(* IEC 61131-3 sources: plc-st-coding-agent/progress/evidence/f14_v6_public_pilot_20261112/jobs/custom_minimax-m27, 44 files *)

(* ---- public-easy-01.candidate_01.st ---- *)
FUNCTION_BLOCK FillLineControl
VAR_INPUT
    bottleSensor           : BOOL;
    cleaningConfirmButton  : BOOL;
    fillingConfirmButton   : BOOL;
    cappingConfirmButton   : BOOL;
    packingConfirmButton   : BOOL;
    finishedButton         : BOOL;
END_VAR

VAR_OUTPUT
    Pump_Motor         : BOOL;
    Filling_Valve      : BOOL;
    Capping_Machine    : BOOL;
    Packing_Machine    : BOOL;
    Completion_Light   : BOOL;
END_VAR

VAR
    eState : INT;
    tmp_R_TRIG_cleaning : R_TRIG;
    tmp_R_TRIG_filling  : R_TRIG;
    tmp_R_TRIG_capping  : R_TRIG;
    tmp_R_TRIG_packing  : R_TRIG;
    tmp_R_TRIG_finished : R_TRIG;
END_VAR

VAR CONSTANT
    STATE_IDLE      : INT := 0;
    STATE_CLEANING  : INT := 1;
    STATE_FILLING   : INT := 2;
    STATE_CAPPING   : INT := 3;
    STATE_PACKING   : INT := 4;
    STATE_COMPLETED : INT := 5;
END_VAR

(* ENGINEERING_CONTRACT
  State machine for automated filling line (6 states, linear sequence):
  +------------------+-------------------------------+-------------------+-------------------+---------------------------+
  | State            | Active Outputs                | Retention         | Deactivation      | Trigger                   |
  +------------------+-------------------------------+-------------------+-------------------+---------------------------+
  | IDLE (0)         | none                          | N/A               | N/A               | bottleSensor=TRUE         |
  | CLEANING (1)     | Pump_Motor=TRUE               | Hold until next   | Next state enter  | cleaningConfirmButton edge|
  | FILLING (2)      | Filling_Valve=TRUE            | Hold until next   | Next state enter  | fillingConfirmButton edge |
  | CAPPING (3)      | Capping_Machine=TRUE          | Hold until next   | Next state enter  | cappingConfirmButton edge |
  | PACKING (4)      | Packing_Machine=TRUE          | Hold until next   | Next state enter  | packingConfirmButton edge |
  | COMPLETED (5)    | Completion_Light=TRUE         | Hold until reset  | finishedButton edge | packingConfirmButton edge|
  +------------------+-------------------------------+-------------------+-------------------+---------------------------+
  Priority: Same-scan parallel evaluation, outputs set per state at scan end.
  References: PUB003(cleaning pump start), PUB004(cleaningConfirmButton),
              PUB005(fillingConfirmButton), PUB006(cappingConfirmButton),
              PUB007(packingConfirmButton), PUB008(finishedButton reset).
*)
(* CONTRACT_RULES [{"kind":"hold_until_reset","output":"Completion_Light","set_input":"packingConfirmButton","reset_input":"finishedButton"}] *)

tmp_R_TRIG_cleaning(CLK := cleaningConfirmButton);
tmp_R_TRIG_filling(CLK  := fillingConfirmButton);
tmp_R_TRIG_capping(CLK  := cappingConfirmButton);
tmp_R_TRIG_packing(CLK  := packingConfirmButton);
tmp_R_TRIG_finished(CLK := finishedButton);

CASE eState OF
    STATE_IDLE:
        Pump_Motor       := FALSE;
        Filling_Valve    := FALSE;
        Capping_Machine  := FALSE;
        Packing_Machine  := FALSE;
        Completion_Light := FALSE;

        IF bottleSensor THEN
            eState := STATE_CLEANING;
        END_IF;

    STATE_CLEANING:
        Pump_Motor       := TRUE;
        Filling_Valve    := FALSE;
        Capping_Machine  := FALSE;
        Packing_Machine  := FALSE;
        Completion_Light := FALSE;

        IF tmp_R_TRIG_cleaning.Q THEN
            eState := STATE_FILLING;
        END_IF;

    STATE_FILLING:
        Pump_Motor       := FALSE;
        Filling_Valve    := TRUE;
        Capping_Machine  := FALSE;
        Packing_Machine  := FALSE;
        Completion_Light := FALSE;

        IF tmp_R_TRIG_filling.Q THEN
            eState := STATE_CAPPING;
        END_IF;

    STATE_CAPPING:
        Pump_Motor       := FALSE;
        Filling_Valve    := FALSE;
        Capping_Machine  := TRUE;
        Packing_Machine  := FALSE;
        Completion_Light := FALSE;

        IF tmp_R_TRIG_capping.Q THEN
            eState := STATE_PACKING;
        END_IF;

    STATE_PACKING:
        Pump_Motor       := FALSE;
        Filling_Valve    := FALSE;
        Capping_Machine  := FALSE;
        Packing_Machine  := TRUE;
        Completion_Light := FALSE;

        IF tmp_R_TRIG_packing.Q THEN
            eState := STATE_COMPLETED;
        END_IF;

    STATE_COMPLETED:
        Pump_Motor       := FALSE;
        Filling_Valve    := FALSE;
        Capping_Machine  := FALSE;
        Packing_Machine  := FALSE;
        Completion_Light := TRUE;

        IF tmp_R_TRIG_finished.Q THEN
            eState := STATE_IDLE;
        END_IF;
END_CASE;

END_FUNCTION_BLOCK

(* ---- public-easy-01.candidate_02.st ---- *)
FUNCTION_BLOCK FillLineControl
VAR_INPUT
    bottleSensor           : BOOL;
    cleaningConfirmButton  : BOOL;
    fillingConfirmButton   : BOOL;
    cappingConfirmButton   : BOOL;
    packingConfirmButton   : BOOL;
    finishedButton         : BOOL;
END_VAR

VAR_OUTPUT
    Pump_Motor         : BOOL;
    Filling_Valve      : BOOL;
    Capping_Machine    : BOOL;
    Packing_Machine    : BOOL;
    Completion_Light   : BOOL;
END_VAR

VAR
    eState : INT;
    tmp_R_TRIG_cleaning : R_TRIG;
    tmp_R_TRIG_filling  : R_TRIG;
    tmp_R_TRIG_capping  : R_TRIG;
    tmp_R_TRIG_packing  : R_TRIG;
    tmp_R_TRIG_finished : R_TRIG;
END_VAR

VAR CONSTANT
    STATE_IDLE      : INT := 0;
    STATE_CLEANING  : INT := 1;
    STATE_FILLING   : INT := 2;
    STATE_CAPPING   : INT := 3;
    STATE_PACKING   : INT := 4;
    STATE_COMPLETED : INT := 5;
END_VAR

(* ENGINEERING_CONTRACT
  State machine for automated filling line (6 states, linear sequence):
  +------------------+-------------------------------+-------------------+-------------------+---------------------------+
  | State            | Active Outputs                | Retention         | Deactivation      | Trigger                   |
  +------------------+-------------------------------+-------------------+-------------------+---------------------------+
  | IDLE (0)         | none                          | N/A               | N/A               | bottleSensor=TRUE         |
  | CLEANING (1)     | Pump_Motor=TRUE               | Hold until next   | Next state enter  | cleaningConfirmButton edge|
  | FILLING (2)      | Filling_Valve=TRUE            | Hold until next   | Next state enter  | fillingConfirmButton edge |
  | CAPPING (3)      | Capping_Machine=TRUE          | Hold until next   | Next state enter  | cappingConfirmButton edge |
  | PACKING (4)      | Packing_Machine=TRUE          | Hold until next   | Next state enter  | packingConfirmButton edge |
  | COMPLETED (5)    | Completion_Light=TRUE         | Hold until reset  | finishedButton edge | -                      |
  +------------------+-------------------------------+-------------------+-------------------+---------------------------+
  Priority: Same-scan parallel evaluation, outputs set per state at scan end.
  Completion_Light set_input (packingConfirmButton) requires reaching STATE_PACKING first;
  this prerequisite cannot be expressed in flat contract format and is handled by the
  state machine logic. PUB003-PUB008 define all transitions.
*)
(* CONTRACT_RULES [] *)

tmp_R_TRIG_cleaning(CLK := cleaningConfirmButton);
tmp_R_TRIG_filling(CLK  := fillingConfirmButton);
tmp_R_TRIG_capping(CLK  := cappingConfirmButton);
tmp_R_TRIG_packing(CLK  := packingConfirmButton);
tmp_R_TRIG_finished(CLK := finishedButton);

CASE eState OF
    STATE_IDLE:
        Pump_Motor       := FALSE;
        Filling_Valve    := FALSE;
        Capping_Machine  := FALSE;
        Packing_Machine  := FALSE;
        Completion_Light := FALSE;

        IF bottleSensor THEN
            eState := STATE_CLEANING;
        END_IF;

    STATE_CLEANING:
        Pump_Motor       := TRUE;
        Filling_Valve    := FALSE;
        Capping_Machine  := FALSE;
        Packing_Machine  := FALSE;
        Completion_Light := FALSE;

        IF tmp_R_TRIG_cleaning.Q THEN
            eState := STATE_FILLING;
        END_IF;

    STATE_FILLING:
        Pump_Motor       := FALSE;
        Filling_Valve    := TRUE;
        Capping_Machine  := FALSE;
        Packing_Machine  := FALSE;
        Completion_Light := FALSE;

        IF tmp_R_TRIG_filling.Q THEN
            eState := STATE_CAPPING;
        END_IF;

    STATE_CAPPING:
        Pump_Motor       := FALSE;
        Filling_Valve    := FALSE;
        Capping_Machine  := TRUE;
        Packing_Machine  := FALSE;
        Completion_Light := FALSE;

        IF tmp_R_TRIG_capping.Q THEN
            eState := STATE_PACKING;
        END_IF;

    STATE_PACKING:
        Pump_Motor       := FALSE;
        Filling_Valve    := FALSE;
        Capping_Machine  := FALSE;
        Packing_Machine  := TRUE;
        Completion_Light := FALSE;

        IF tmp_R_TRIG_packing.Q THEN
            eState := STATE_COMPLETED;
        END_IF;

    STATE_COMPLETED:
        Pump_Motor       := FALSE;
        Filling_Valve    := FALSE;
        Capping_Machine  := FALSE;
        Packing_Machine  := FALSE;
        Completion_Light := TRUE;

        IF tmp_R_TRIG_finished.Q THEN
            eState := STATE_IDLE;
        END_IF;
END_CASE;

END_FUNCTION_BLOCK

(* ---- public-easy-01.candidate_03.st ---- *)
FUNCTION_BLOCK FillLineControl
VAR_INPUT
    bottleSensor           : BOOL;
    cleaningConfirmButton  : BOOL;
    fillingConfirmButton   : BOOL;
    cappingConfirmButton   : BOOL;
    packingConfirmButton   : BOOL;
    finishedButton         : BOOL;
END_VAR

VAR_OUTPUT
    Pump_Motor         : BOOL;
    Filling_Valve      : BOOL;
    Capping_Machine    : BOOL;
    Packing_Machine    : BOOL;
    Completion_Light   : BOOL;
END_VAR

VAR
    eState : INT;
    tmp_R_TRIG_cleaning : R_TRIG;
    tmp_R_TRIG_filling  : R_TRIG;
    tmp_R_TRIG_capping  : R_TRIG;
    tmp_R_TRIG_packing  : R_TRIG;
    tmp_R_TRIG_finished : R_TRIG;
END_VAR

VAR CONSTANT
    STATE_IDLE      : INT := 0;
    STATE_CLEANING  : INT := 1;
    STATE_FILLING   : INT := 2;
    STATE_CAPPING   : INT := 3;
    STATE_PACKING   : INT := 4;
END_VAR

(* ENGINEERING_CONTRACT
  State machine for automated filling line (5 states, linear sequence):
  +------------------+-------------------------------+-------------------+-------------------+---------------------------+
  | State            | Active Outputs                | Retention         | Deactivation      | Trigger                   |
  +------------------+-------------------------------+-------------------+-------------------+---------------------------+
  | IDLE (0)         | none                          | N/A               | N/A               | bottleSensor=TRUE         |
  | CLEANING (1)     | Pump_Motor=TRUE               | Hold until next   | Next state enter  | cleaningConfirmButton edge|
  | FILLING (2)      | Filling_Valve=TRUE            | Hold until next   | Next state enter  | fillingConfirmButton edge |
  | CAPPING (3)      | Capping_Machine=TRUE          | Hold until next   | Next state enter  | cappingConfirmButton edge |
  | PACKING (4)      | Packing_Machine=TRUE          | Hold until next   | Next state enter  | packingConfirmButton edge |
  +------------------+-------------------------------+-------------------+-------------------+---------------------------+
  Completion_Light: PUB007 latched output, set by packingConfirmButton edge,
                    reset by finishedButton edge. Independent of state machine.
  Priority: Same-scan parallel evaluation, outputs set per state at scan end.
  References: PUB003(cleaning pump start), PUB004(cleaningConfirmButton),
              PUB005(fillingConfirmButton), PUB006(cappingConfirmButton),
              PUB007(packingConfirmButton triggers Completion_Light),
              PUB008(finishedButton reset).
*)
(* CONTRACT_RULES [{"kind":"hold_until_reset","output":"Completion_Light","set_input":"packingConfirmButton","reset_input":"finishedButton"}] *)

tmp_R_TRIG_cleaning(CLK := cleaningConfirmButton);
tmp_R_TRIG_filling(CLK  := fillingConfirmButton);
tmp_R_TRIG_capping(CLK  := cappingConfirmButton);
tmp_R_TRIG_packing(CLK  := packingConfirmButton);
tmp_R_TRIG_finished(CLK := finishedButton);

CASE eState OF
    STATE_IDLE:
        Pump_Motor       := FALSE;
        Filling_Valve    := FALSE;
        Capping_Machine  := FALSE;
        Packing_Machine  := FALSE;

        IF bottleSensor THEN
            eState := STATE_CLEANING;
        END_IF;

    STATE_CLEANING:
        Pump_Motor       := TRUE;
        Filling_Valve    := FALSE;
        Capping_Machine  := FALSE;
        Packing_Machine  := FALSE;

        IF tmp_R_TRIG_cleaning.Q THEN
            eState := STATE_FILLING;
        END_IF;

    STATE_FILLING:
        Pump_Motor       := FALSE;
        Filling_Valve    := TRUE;
        Capping_Machine  := FALSE;
        Packing_Machine  := FALSE;

        IF tmp_R_TRIG_filling.Q THEN
            eState := STATE_CAPPING;
        END_IF;

    STATE_CAPPING:
        Pump_Motor       := FALSE;
        Filling_Valve    := FALSE;
        Capping_Machine  := TRUE;
        Packing_Machine  := FALSE;

        IF tmp_R_TRIG_capping.Q THEN
            eState := STATE_PACKING;
        END_IF;

    STATE_PACKING:
        Pump_Motor       := FALSE;
        Filling_Valve    := FALSE;
        Capping_Machine  := FALSE;
        Packing_Machine  := TRUE;

        IF tmp_R_TRIG_packing.Q THEN
            eState := STATE_IDLE;
        END_IF;
END_CASE;

IF tmp_R_TRIG_packing.Q THEN
    Completion_Light := TRUE;
END_IF;

IF tmp_R_TRIG_finished.Q THEN
    Completion_Light := FALSE;
END_IF;

END_FUNCTION_BLOCK

(* ---- public-easy-01.candidate_04.st ---- *)
FUNCTION_BLOCK FillLineControl
VAR_INPUT
    bottleSensor           : BOOL;
    cleaningConfirmButton  : BOOL;
    fillingConfirmButton   : BOOL;
    cappingConfirmButton   : BOOL;
    packingConfirmButton   : BOOL;
    finishedButton         : BOOL;
END_VAR

VAR_OUTPUT
    Pump_Motor         : BOOL;
    Filling_Valve      : BOOL;
    Capping_Machine    : BOOL;
    Packing_Machine    : BOOL;
    Completion_Light   : BOOL;
END_VAR

VAR
    eState : INT := 0;
END_VAR

VAR CONSTANT
    STATE_IDLE      : INT := 0;
    STATE_CLEANING  : INT := 1;
    STATE_FILLING   : INT := 2;
    STATE_CAPPING   : INT := 3;
    STATE_PACKING   : INT := 4;
    STATE_COMPLETED : INT := 5;
END_VAR

(* ENGINEERING_CONTRACT
  Linear 6-state filling line with sequential transitions:
  +------------------+-------------------------------+-------------------+-------------------+---------------------------+
  | State            | Active Outputs                | Retention         | Deactivation      | Trigger                   |
  +------------------+-------------------------------+-------------------+-------------------+---------------------------+
  | IDLE (0)         | none                          | N/A               | N/A               | bottleSensor=TRUE         |
  | CLEANING (1)     | Pump_Motor=TRUE               | Hold until next   | Next state enter  | cleaningConfirmButton=TRUE|
  | FILLING (2)      | Filling_Valve=TRUE            | Hold until next   | Next state enter  | fillingConfirmButton=TRUE |
  | CAPPING (3)      | Capping_Machine=TRUE          | Hold until next   | Next state enter  | cappingConfirmButton=TRUE |
  | PACKING (4)      | Packing_Machine=TRUE          | Hold until next   | Next state enter  | packingConfirmButton=TRUE |
  | COMPLETED (5)    | Completion_Light=TRUE         | Hold until reset  | finishedButton=TRUE | packingConfirmButton=TRUE|
  +------------------+-------------------------------+-------------------+-------------------+---------------------------+
  Priority: Outputs set immediately on state entry before transition checks.
  References: PUB003(cleaning pump), PUB004(cleaningConfirmButton),
              PUB005(fillingConfirmButton), PUB006(cappingConfirmButton),
              PUB007(packingConfirmButton), PUB008(finishedButton reset).
*)
(* CONTRACT_RULES [{"kind":"hold_until_reset","output":"Completion_Light","set_input":"packingConfirmButton","reset_input":"finishedButton"}] *)

CASE eState OF
    STATE_IDLE:
        IF bottleSensor THEN
            eState := STATE_CLEANING;
        END_IF;

    STATE_CLEANING:
        IF cleaningConfirmButton THEN
            eState := STATE_FILLING;
        END_IF;

    STATE_FILLING:
        IF fillingConfirmButton THEN
            eState := STATE_CAPPING;
        END_IF;

    STATE_CAPPING:
        IF cappingConfirmButton THEN
            eState := STATE_PACKING;
        END_IF;

    STATE_PACKING:
        IF packingConfirmButton THEN
            eState := STATE_COMPLETED;
        END_IF;

    STATE_COMPLETED:
        IF finishedButton THEN
            eState := STATE_IDLE;
        END_IF;
END_CASE;

Pump_Motor       := (eState = STATE_CLEANING);
Filling_Valve    := (eState = STATE_FILLING);
Capping_Machine  := (eState = STATE_CAPPING);
Packing_Machine  := (eState = STATE_PACKING);
Completion_Light := (eState = STATE_COMPLETED);

END_FUNCTION_BLOCK

(* ---- public-easy-01.raw_candidate_01.st ---- *)
FUNCTION_BLOCK FillLineControl
VAR_INPUT
    bottleSensor           : BOOL;
    cleaningConfirmButton  : BOOL;
    fillingConfirmButton   : BOOL;
    cappingConfirmButton   : BOOL;
    packingConfirmButton   : BOOL;
    finishedButton         : BOOL;
END_VAR

VAR_OUTPUT
    Pump_Motor         : BOOL;
    Filling_Valve      : BOOL;
    Capping_Machine    : BOOL;
    Packing_Machine    : BOOL;
    Completion_Light   : BOOL;
END_VAR

VAR
    eState : INT;
    tmp_R_TRIG_cleaning : R_TRIG;
    tmp_R_TRIG_filling  : R_TRIG;
    tmp_R_TRIG_capping  : R_TRIG;
    tmp_R_TRIG_packing  : R_TRIG;
    tmp_R_TRIG_finished : R_TRIG;
END_VAR

VAR CONSTANT
    STATE_IDLE      : INT := 0;
    STATE_CLEANING  : INT := 1;
    STATE_FILLING   : INT := 2;
    STATE_CAPPING   : INT := 3;
    STATE_PACKING   : INT := 4;
    STATE_COMPLETED : INT := 5;
END_VAR

(* ENGINEERING_CONTRACT
  State machine for automated filling line (6 states, linear sequence):
  +------------------+-------------------------------+-------------------+-------------------+---------------------------+
  | State            | Active Outputs                | Retention         | Deactivation      | Trigger                   |
  +------------------+-------------------------------+-------------------+-------------------+---------------------------+
  | IDLE (0)         | none                          | N/A               | N/A               | bottleSensor=TRUE         |
  | CLEANING (1)     | Pump_Motor=TRUE               | Hold until next   | Next state enter  | cleaningConfirmButton edge|
  | FILLING (2)      | Filling_Valve=TRUE            | Hold until next   | Next state enter  | fillingConfirmButton edge |
  | CAPPING (3)      | Capping_Machine=TRUE          | Hold until next   | Next state enter  | cappingConfirmButton edge |
  | PACKING (4)      | Packing_Machine=TRUE          | Hold until next   | Next state enter  | packingConfirmButton edge |
  | COMPLETED (5)    | Completion_Light=TRUE         | Hold until reset  | finishedButton edge | packingConfirmButton edge|
  +------------------+-------------------------------+-------------------+-------------------+---------------------------+
  Priority: Same-scan parallel evaluation, outputs set per state at scan end.
  References: PUB003(cleaning pump start), PUB004(cleaningConfirmButton),
              PUB005(fillingConfirmButton), PUB006(cappingConfirmButton),
              PUB007(packingConfirmButton), PUB008(finishedButton reset).
*)
(* CONTRACT_RULES [{"kind":"hold_until_reset","output":"Completion_Light","set_input":"packingConfirmButton","reset_input":"finishedButton"}] *)

tmp_R_TRIG_cleaning(CLK := cleaningConfirmButton);
tmp_R_TRIG_filling(CLK  := fillingConfirmButton);
tmp_R_TRIG_capping(CLK  := cappingConfirmButton);
tmp_R_TRIG_packing(CLK  := packingConfirmButton);
tmp_R_TRIG_finished(CLK := finishedButton);

CASE eState OF
    STATE_IDLE:
        Pump_Motor       := FALSE;
        Filling_Valve    := FALSE;
        Capping_Machine  := FALSE;
        Packing_Machine  := FALSE;
        Completion_Light := FALSE;

        IF bottleSensor THEN
            eState := STATE_CLEANING;
        END_IF;

    STATE_CLEANING:
        Pump_Motor       := TRUE;
        Filling_Valve    := FALSE;
        Capping_Machine  := FALSE;
        Packing_Machine  := FALSE;
        Completion_Light := FALSE;

        IF tmp_R_TRIG_cleaning.Q THEN
            eState := STATE_FILLING;
        END_IF;

    STATE_FILLING:
        Pump_Motor       := FALSE;
        Filling_Valve    := TRUE;
        Capping_Machine  := FALSE;
        Packing_Machine  := FALSE;
        Completion_Light := FALSE;

        IF tmp_R_TRIG_filling.Q THEN
            eState := STATE_CAPPING;
        END_IF;

    STATE_CAPPING:
        Pump_Motor       := FALSE;
        Filling_Valve    := FALSE;
        Capping_Machine  := TRUE;
        Packing_Machine  := FALSE;
        Completion_Light := FALSE;

        IF tmp_R_TRIG_capping.Q THEN
            eState := STATE_PACKING;
        END_IF;

    STATE_PACKING:
        Pump_Motor       := FALSE;
        Filling_Valve    := FALSE;
        Capping_Machine  := FALSE;
        Packing_Machine  := TRUE;
        Completion_Light := FALSE;

        IF tmp_R_TRIG_packing.Q THEN
            eState := STATE_COMPLETED;
        END_IF;

    STATE_COMPLETED:
        Pump_Motor       := FALSE;
        Filling_Valve    := FALSE;
        Capping_Machine  := FALSE;
        Packing_Machine  := FALSE;
        Completion_Light := TRUE;

        IF tmp_R_TRIG_finished.Q THEN
            eState := STATE_IDLE;
        END_IF;
END_CASE;

END_FUNCTION_BLOCK

(* ---- public-easy-01.raw_candidate_02.st ---- *)
FUNCTION_BLOCK FillLineControl
VAR_INPUT
    bottleSensor           : BOOL;
    cleaningConfirmButton  : BOOL;
    fillingConfirmButton   : BOOL;
    cappingConfirmButton   : BOOL;
    packingConfirmButton   : BOOL;
    finishedButton         : BOOL;
END_VAR

VAR_OUTPUT
    Pump_Motor         : BOOL;
    Filling_Valve      : BOOL;
    Capping_Machine    : BOOL;
    Packing_Machine    : BOOL;
    Completion_Light   : BOOL;
END_VAR

VAR
    eState : INT;
    tmp_R_TRIG_cleaning : R_TRIG;
    tmp_R_TRIG_filling  : R_TRIG;
    tmp_R_TRIG_capping  : R_TRIG;
    tmp_R_TRIG_packing  : R_TRIG;
    tmp_R_TRIG_finished : R_TRIG;
END_VAR

VAR CONSTANT
    STATE_IDLE      : INT := 0;
    STATE_CLEANING  : INT := 1;
    STATE_FILLING   : INT := 2;
    STATE_CAPPING   : INT := 3;
    STATE_PACKING   : INT := 4;
    STATE_COMPLETED : INT := 5;
END_VAR

(* ENGINEERING_CONTRACT
  State machine for automated filling line (6 states, linear sequence):
  +------------------+-------------------------------+-------------------+-------------------+---------------------------+
  | State            | Active Outputs                | Retention         | Deactivation      | Trigger                   |
  +------------------+-------------------------------+-------------------+-------------------+---------------------------+
  | IDLE (0)         | none                          | N/A               | N/A               | bottleSensor=TRUE         |
  | CLEANING (1)     | Pump_Motor=TRUE               | Hold until next   | Next state enter  | cleaningConfirmButton edge|
  | FILLING (2)      | Filling_Valve=TRUE            | Hold until next   | Next state enter  | fillingConfirmButton edge |
  | CAPPING (3)      | Capping_Machine=TRUE          | Hold until next   | Next state enter  | cappingConfirmButton edge |
  | PACKING (4)      | Packing_Machine=TRUE          | Hold until next   | Next state enter  | packingConfirmButton edge |
  | COMPLETED (5)    | Completion_Light=TRUE         | Hold until reset  | finishedButton edge | -                      |
  +------------------+-------------------------------+-------------------+-------------------+---------------------------+
  Priority: Same-scan parallel evaluation, outputs set per state at scan end.
  Completion_Light set_input (packingConfirmButton) requires reaching STATE_PACKING first;
  this prerequisite cannot be expressed in flat contract format and is handled by the
  state machine logic. PUB003-PUB008 define all transitions.
*)
(* CONTRACT_RULES [] *)

tmp_R_TRIG_cleaning(CLK := cleaningConfirmButton);
tmp_R_TRIG_filling(CLK  := fillingConfirmButton);
tmp_R_TRIG_capping(CLK  := cappingConfirmButton);
tmp_R_TRIG_packing(CLK  := packingConfirmButton);
tmp_R_TRIG_finished(CLK := finishedButton);

CASE eState OF
    STATE_IDLE:
        Pump_Motor       := FALSE;
        Filling_Valve    := FALSE;
        Capping_Machine  := FALSE;
        Packing_Machine  := FALSE;
        Completion_Light := FALSE;

        IF bottleSensor THEN
            eState := STATE_CLEANING;
        END_IF;

    STATE_CLEANING:
        Pump_Motor       := TRUE;
        Filling_Valve    := FALSE;
        Capping_Machine  := FALSE;
        Packing_Machine  := FALSE;
        Completion_Light := FALSE;

        IF tmp_R_TRIG_cleaning.Q THEN
            eState := STATE_FILLING;
        END_IF;

    STATE_FILLING:
        Pump_Motor       := FALSE;
        Filling_Valve    := TRUE;
        Capping_Machine  := FALSE;
        Packing_Machine  := FALSE;
        Completion_Light := FALSE;

        IF tmp_R_TRIG_filling.Q THEN
            eState := STATE_CAPPING;
        END_IF;

    STATE_CAPPING:
        Pump_Motor       := FALSE;
        Filling_Valve    := FALSE;
        Capping_Machine  := TRUE;
        Packing_Machine  := FALSE;
        Completion_Light := FALSE;

        IF tmp_R_TRIG_capping.Q THEN
            eState := STATE_PACKING;
        END_IF;

    STATE_PACKING:
        Pump_Motor       := FALSE;
        Filling_Valve    := FALSE;
        Capping_Machine  := FALSE;
        Packing_Machine  := TRUE;
        Completion_Light := FALSE;

        IF tmp_R_TRIG_packing.Q THEN
            eState := STATE_COMPLETED;
        END_IF;

    STATE_COMPLETED:
        Pump_Motor       := FALSE;
        Filling_Valve    := FALSE;
        Capping_Machine  := FALSE;
        Packing_Machine  := FALSE;
        Completion_Light := TRUE;

        IF tmp_R_TRIG_finished.Q THEN
            eState := STATE_IDLE;
        END_IF;
END_CASE;

END_FUNCTION_BLOCK

(* ---- public-easy-01.raw_candidate_03.st ---- *)
FUNCTION_BLOCK FillLineControl
VAR_INPUT
    bottleSensor           : BOOL;
    cleaningConfirmButton  : BOOL;
    fillingConfirmButton   : BOOL;
    cappingConfirmButton   : BOOL;
    packingConfirmButton   : BOOL;
    finishedButton         : BOOL;
END_VAR

VAR_OUTPUT
    Pump_Motor         : BOOL;
    Filling_Valve      : BOOL;
    Capping_Machine    : BOOL;
    Packing_Machine    : BOOL;
    Completion_Light   : BOOL;
END_VAR

VAR
    eState : INT;
    tmp_R_TRIG_cleaning : R_TRIG;
    tmp_R_TRIG_filling  : R_TRIG;
    tmp_R_TRIG_capping  : R_TRIG;
    tmp_R_TRIG_packing  : R_TRIG;
    tmp_R_TRIG_finished : R_TRIG;
END_VAR

VAR CONSTANT
    STATE_IDLE      : INT := 0;
    STATE_CLEANING  : INT := 1;
    STATE_FILLING   : INT := 2;
    STATE_CAPPING   : INT := 3;
    STATE_PACKING   : INT := 4;
END_VAR

(* ENGINEERING_CONTRACT
  State machine for automated filling line (5 states, linear sequence):
  +------------------+-------------------------------+-------------------+-------------------+---------------------------+
  | State            | Active Outputs                | Retention         | Deactivation      | Trigger                   |
  +------------------+-------------------------------+-------------------+-------------------+---------------------------+
  | IDLE (0)         | none                          | N/A               | N/A               | bottleSensor=TRUE         |
  | CLEANING (1)     | Pump_Motor=TRUE               | Hold until next   | Next state enter  | cleaningConfirmButton edge|
  | FILLING (2)      | Filling_Valve=TRUE            | Hold until next   | Next state enter  | fillingConfirmButton edge |
  | CAPPING (3)      | Capping_Machine=TRUE          | Hold until next   | Next state enter  | cappingConfirmButton edge |
  | PACKING (4)      | Packing_Machine=TRUE          | Hold until next   | Next state enter  | packingConfirmButton edge |
  +------------------+-------------------------------+-------------------+-------------------+---------------------------+
  Completion_Light: PUB007 latched output, set by packingConfirmButton edge,
                    reset by finishedButton edge. Independent of state machine.
  Priority: Same-scan parallel evaluation, outputs set per state at scan end.
  References: PUB003(cleaning pump start), PUB004(cleaningConfirmButton),
              PUB005(fillingConfirmButton), PUB006(cappingConfirmButton),
              PUB007(packingConfirmButton triggers Completion_Light),
              PUB008(finishedButton reset).
*)
(* CONTRACT_RULES [{"kind":"hold_until_reset","output":"Completion_Light","set_input":"packingConfirmButton","reset_input":"finishedButton"}] *)

tmp_R_TRIG_cleaning(CLK := cleaningConfirmButton);
tmp_R_TRIG_filling(CLK  := fillingConfirmButton);
tmp_R_TRIG_capping(CLK  := cappingConfirmButton);
tmp_R_TRIG_packing(CLK  := packingConfirmButton);
tmp_R_TRIG_finished(CLK := finishedButton);

CASE eState OF
    STATE_IDLE:
        Pump_Motor       := FALSE;
        Filling_Valve    := FALSE;
        Capping_Machine  := FALSE;
        Packing_Machine  := FALSE;

        IF bottleSensor THEN
            eState := STATE_CLEANING;
        END_IF;

    STATE_CLEANING:
        Pump_Motor       := TRUE;
        Filling_Valve    := FALSE;
        Capping_Machine  := FALSE;
        Packing_Machine  := FALSE;

        IF tmp_R_TRIG_cleaning.Q THEN
            eState := STATE_FILLING;
        END_IF;

    STATE_FILLING:
        Pump_Motor       := FALSE;
        Filling_Valve    := TRUE;
        Capping_Machine  := FALSE;
        Packing_Machine  := FALSE;

        IF tmp_R_TRIG_filling.Q THEN
            eState := STATE_CAPPING;
        END_IF;

    STATE_CAPPING:
        Pump_Motor       := FALSE;
        Filling_Valve    := FALSE;
        Capping_Machine  := TRUE;
        Packing_Machine  := FALSE;

        IF tmp_R_TRIG_capping.Q THEN
            eState := STATE_PACKING;
        END_IF;

    STATE_PACKING:
        Pump_Motor       := FALSE;
        Filling_Valve    := FALSE;
        Capping_Machine  := FALSE;
        Packing_Machine  := TRUE;

        IF tmp_R_TRIG_packing.Q THEN
            eState := STATE_IDLE;
        END_IF;
END_CASE;

IF tmp_R_TRIG_packing.Q THEN
    Completion_Light := TRUE;
END_IF;

IF tmp_R_TRIG_finished.Q THEN
    Completion_Light := FALSE;
END_IF;

END_FUNCTION_BLOCK

(* ---- public-easy-01.raw_candidate_04.st ---- *)
FUNCTION_BLOCK FillLineControl
VAR_INPUT
    bottleSensor           : BOOL;
    cleaningConfirmButton  : BOOL;
    fillingConfirmButton   : BOOL;
    cappingConfirmButton   : BOOL;
    packingConfirmButton   : BOOL;
    finishedButton         : BOOL;
END_VAR

VAR_OUTPUT
    Pump_Motor         : BOOL;
    Filling_Valve      : BOOL;
    Capping_Machine    : BOOL;
    Packing_Machine    : BOOL;
    Completion_Light   : BOOL;
END_VAR

VAR
    eState : INT := 0;
END_VAR

VAR CONSTANT
    STATE_IDLE      : INT := 0;
    STATE_CLEANING  : INT := 1;
    STATE_FILLING   : INT := 2;
    STATE_CAPPING   : INT := 3;
    STATE_PACKING   : INT := 4;
    STATE_COMPLETED : INT := 5;
END_VAR

(* ENGINEERING_CONTRACT
  Linear 6-state filling line with sequential transitions:
  +------------------+-------------------------------+-------------------+-------------------+---------------------------+
  | State            | Active Outputs                | Retention         | Deactivation      | Trigger                   |
  +------------------+-------------------------------+-------------------+-------------------+---------------------------+
  | IDLE (0)         | none                          | N/A               | N/A               | bottleSensor=TRUE         |
  | CLEANING (1)     | Pump_Motor=TRUE               | Hold until next   | Next state enter  | cleaningConfirmButton=TRUE|
  | FILLING (2)      | Filling_Valve=TRUE            | Hold until next   | Next state enter  | fillingConfirmButton=TRUE |
  | CAPPING (3)      | Capping_Machine=TRUE          | Hold until next   | Next state enter  | cappingConfirmButton=TRUE |
  | PACKING (4)      | Packing_Machine=TRUE          | Hold until next   | Next state enter  | packingConfirmButton=TRUE |
  | COMPLETED (5)    | Completion_Light=TRUE         | Hold until reset  | finishedButton=TRUE | packingConfirmButton=TRUE|
  +------------------+-------------------------------+-------------------+-------------------+---------------------------+
  Priority: Outputs set immediately on state entry before transition checks.
  References: PUB003(cleaning pump), PUB004(cleaningConfirmButton),
              PUB005(fillingConfirmButton), PUB006(cappingConfirmButton),
              PUB007(packingConfirmButton), PUB008(finishedButton reset).
*)
(* CONTRACT_RULES [{"kind":"hold_until_reset","output":"Completion_Light","set_input":"packingConfirmButton","reset_input":"finishedButton"}] *)

CASE eState OF
    STATE_IDLE:
        IF bottleSensor THEN
            eState := STATE_CLEANING;
        END_IF;

    STATE_CLEANING:
        IF cleaningConfirmButton THEN
            eState := STATE_FILLING;
        END_IF;

    STATE_FILLING:
        IF fillingConfirmButton THEN
            eState := STATE_CAPPING;
        END_IF;

    STATE_CAPPING:
        IF cappingConfirmButton THEN
            eState := STATE_PACKING;
        END_IF;

    STATE_PACKING:
        IF packingConfirmButton THEN
            eState := STATE_COMPLETED;
        END_IF;

    STATE_COMPLETED:
        IF finishedButton THEN
            eState := STATE_IDLE;
        END_IF;
END_CASE;

Pump_Motor       := (eState = STATE_CLEANING);
Filling_Valve    := (eState = STATE_FILLING);
Capping_Machine  := (eState = STATE_CAPPING);
Packing_Machine  := (eState = STATE_PACKING);
Completion_Light := (eState = STATE_COMPLETED);

END_FUNCTION_BLOCK

(* ---- public-easy-04.candidate_01.st ---- *)
FUNCTION_BLOCK FB_JamPumpControl
VAR_INPUT
    VISCOSITY_OK    : BOOL;
    PASTE_E_STOP_NC : BOOL;
    DebounceTime    : TIME;
    CycleTime       : TIME;
END_VAR
VAR_OUTPUT
    VFD_RUN          : BOOL;
    PUMP_MAINT_DUE   : BOOL;
    PUMP_RUNTIME_ACC : LTIME;
END_VAR
VAR
    ViscosityValid : BOOL := FALSE;
    DebounceTimer  : TON;
    tmp_MaintThreshold : LTIME := LTIME#500h;
END_VAR

(* CONTRACT_RULES [] *)

(* ENGINEERING_CONTRACT
+====================+================+==========+=========================+================+===============+
| Output/State       | Activation     | Retention| Reset/Deactivation      | Same-Scan Prio | Boundaries    |
+====================+================+==========+=========================+================+===============+
| VFD_RUN            | ESTOP=TRUE     | Hold     | Immediately on ESTOP=FALSE per PUB003 | Immediate disable | Boolean       |
|                    | AND            |          | No delay on ESTOP loss   |               |               |
|                    | ViscosityValid |          |                          |               |               |
+--------------------+----------------+----------+-------------------------+----------------+---------------+
| ViscosityValid     | TON.Q=TRUE     | Hold TRUE| Invalidate on           | Immediate      | Internal state|
| (internal)         | after          | while    | VISCOSITY_OK=FALSE      | invalidation   |               |
|                    | DebounceTime   | VISCOSITY_OK=TRUE        | per PUB002     |               |               |
+--------------------+----------------+----------+-------------------------+----------------+---------------+
| PUMP_RUNTIME_ACC   | +CycleTime     | Preserve | Only via power-up init  | Increment per  | LTIME, max    |
|                    | per scan while | when     | (PUB006). No auto-reset | scan when      | 500h threshold|
|                    | VFD_RUN=TRUE   | stopped  | specified.              | VFD_RUN=TRUE   | for PUMP_MAINT|
+--------------------+----------------+----------+-------------------------+----------------+---------------+
| PUMP_MAINT_DUE     | Set when       | Hold TRUE| Not specified (informational per PUB005) | At threshold | Boolean       |
|                    | ACC >= 500h    |          | No reset required       |               |               |
+--------------------+----------------+----------+-------------------------+----------------+---------------+
| DebounceTimer      | Start when     | Running  | Reset (ET=TRUE) on      | Clear on input | TON; PT=DebounceTime |
|                    | VISCOSITY_OK   | if input | VISCOSITY_OK=FALSE per  | drop (PUB002)  |               |
|                    | becomes TRUE   | stays TRUE| PUB002                 |               |               |
+--------------------+----------------+----------+-------------------------+----------------+---------------+
*)

CASE BOOL_TO_INT(PASTE_E_STOP_NC) OF
    0: // Emergency stop active
        VFD_RUN := FALSE;
        ViscosityValid := FALSE;
        DebounceTimer(IN := FALSE, PT := DebounceTime);

    1: // Emergency stop cleared - normal operation
        IF NOT VISCOSITY_OK THEN
            ViscosityValid := FALSE;
            DebounceTimer(IN := FALSE, PT := DebounceTime);
        ELSE
            DebounceTimer(IN := TRUE, PT := DebounceTime);
            ViscosityValid := DebounceTimer.Q;
        END_IF;

        VFD_RUN := ViscosityValid;
END_CASE;

IF VFD_RUN THEN
    PUMP_RUNTIME_ACC := PUMP_RUNTIME_ACC + LTIME(CycleTime);
END_IF;

IF PUMP_RUNTIME_ACC >= tmp_MaintThreshold THEN
    PUMP_MAINT_DUE := TRUE;
END_IF;

END_FUNCTION_BLOCK

(* ---- public-easy-04.candidate_02.st ---- *)
FUNCTION_BLOCK FB_JamPumpControl
VAR_INPUT
    VISCOSITY_OK    : BOOL;
    PASTE_E_STOP_NC : BOOL;
    DebounceTime    : TIME;
    CycleTime       : TIME;
END_VAR
VAR_OUTPUT
    VFD_RUN          : BOOL;
    PUMP_MAINT_DUE   : BOOL;
    PUMP_RUNTIME_ACC : LTIME;
END_VAR
VAR
    ViscosityValid : BOOL := FALSE;
    DebounceTimer  : TON;
    tmp_MaintThreshold : LTIME := LTIME#500h;
END_VAR

(* CONTRACT_RULES [] *)

(* ENGINEERING_CONTRACT
+====================+================+==========+=========================+================+===============+
| Output/State       | Activation     | Retention| Reset/Deactivation      | Same-Scan Prio | Boundaries    |
+====================+================+==========+=========================+================+===============+
| VFD_RUN            | ESTOP=TRUE     | Hold     | Immediately on ESTOP=FALSE per PUB003 | Immediate disable | Boolean       |
|                    | AND            |          | No delay on ESTOP loss   |               |               |
|                    | ViscosityValid |          |                          |               |               |
+--------------------+----------------+----------+-------------------------+----------------+---------------+
| ViscosityValid     | TON.Q=TRUE     | Hold TRUE| Invalidate on           | Immediate      | Internal state|
| (internal)         | after          | while    | VISCOSITY_OK=FALSE      | invalidation   |               |
|                    | DebounceTime   | VISCOSITY_OK=TRUE        | per PUB002     |               |               |
+--------------------+----------------+----------+-------------------------+----------------+---------------+
| PUMP_RUNTIME_ACC   | +CycleTime     | Preserve | Only via power-up init  | Increment per  | LTIME, max    |
|                    | per scan while | when     | (PUB006). No auto-reset | scan when      | 500h threshold|
|                    | VFD_RUN=TRUE   | stopped  | specified.              | VFD_RUN=TRUE   | for PUMP_MAINT|
+--------------------+----------------+----------+-------------------------+----------------+---------------+
| PUMP_MAINT_DUE     | Set when       | Hold TRUE| Not specified (informational per PUB005) | At threshold | Boolean       |
|                    | ACC >= 500h    |          | No reset required       |               |               |
+--------------------+----------------+----------+-------------------------+----------------+---------------+
| DebounceTimer      | Start when     | Running  | Reset (ET=TRUE) on      | Clear on input | TON; PT=DebounceTime |
|                    | VISCOSITY_OK   | if input | VISCOSITY_OK=FALSE per  | drop (PUB002)  |               |
|                    | becomes TRUE   | stays TRUE| PUB002                 |               |               |
+--------------------+----------------+----------+-------------------------+----------------+---------------+
*)

CASE BOOL_TO_INT(PASTE_E_STOP_NC) OF
    0: // Emergency stop active
        VFD_RUN := FALSE;
        ViscosityValid := FALSE;
        DebounceTimer(IN := FALSE, PT := DebounceTime);

    1: // Emergency stop cleared - normal operation
        IF NOT VISCOSITY_OK THEN
            ViscosityValid := FALSE;
            DebounceTimer(IN := FALSE, PT := DebounceTime);
        ELSE
            DebounceTimer(IN := TRUE, PT := DebounceTime);
            ViscosityValid := DebounceTimer.Q;
        END_IF;

        VFD_RUN := ViscosityValid;
END_CASE;

IF VFD_RUN THEN
    PUMP_RUNTIME_ACC := PUMP_RUNTIME_ACC + TIME_TO_LTIME(CycleTime);
END_IF;

IF PUMP_RUNTIME_ACC >= tmp_MaintThreshold THEN
    PUMP_MAINT_DUE := TRUE;
END_IF;

END_FUNCTION_BLOCK

(* ---- public-easy-04.raw_candidate_01.st ---- *)
FUNCTION_BLOCK FB_JamPumpControl
VAR_INPUT
    VISCOSITY_OK    : BOOL;
    PASTE_E_STOP_NC : BOOL;
    DebounceTime    : TIME;
    CycleTime       : TIME;
END_VAR
VAR_OUTPUT
    VFD_RUN          : BOOL;
    PUMP_MAINT_DUE   : BOOL;
    PUMP_RUNTIME_ACC : LTIME;
END_VAR
VAR
    ViscosityValid : BOOL := FALSE;
    DebounceTimer  : TON;
    tmp_MaintThreshold : LTIME := LTIME#500h;
END_VAR

(* CONTRACT_RULES [] *)

(* ENGINEERING_CONTRACT
+====================+================+==========+=========================+================+===============+
| Output/State       | Activation     | Retention| Reset/Deactivation      | Same-Scan Prio | Boundaries    |
+====================+================+==========+=========================+================+===============+
| VFD_RUN            | ESTOP=TRUE     | Hold     | Immediately on ESTOP=FALSE per PUB003 | Immediate disable | Boolean       |
|                    | AND            |          | No delay on ESTOP loss   |               |               |
|                    | ViscosityValid |          |                          |               |               |
+--------------------+----------------+----------+-------------------------+----------------+---------------+
| ViscosityValid     | TON.Q=TRUE     | Hold TRUE| Invalidate on           | Immediate      | Internal state|
| (internal)         | after          | while    | VISCOSITY_OK=FALSE      | invalidation   |               |
|                    | DebounceTime   | VISCOSITY_OK=TRUE        | per PUB002     |               |               |
+--------------------+----------------+----------+-------------------------+----------------+---------------+
| PUMP_RUNTIME_ACC   | +CycleTime     | Preserve | Only via power-up init  | Increment per  | LTIME, max    |
|                    | per scan while | when     | (PUB006). No auto-reset | scan when      | 500h threshold|
|                    | VFD_RUN=TRUE   | stopped  | specified.              | VFD_RUN=TRUE   | for PUMP_MAINT|
+--------------------+----------------+----------+-------------------------+----------------+---------------+
| PUMP_MAINT_DUE     | Set when       | Hold TRUE| Not specified (informational per PUB005) | At threshold | Boolean       |
|                    | ACC >= 500h    |          | No reset required       |               |               |
+--------------------+----------------+----------+-------------------------+----------------+---------------+
| DebounceTimer      | Start when     | Running  | Reset (ET=TRUE) on      | Clear on input | TON; PT=DebounceTime |
|                    | VISCOSITY_OK   | if input | VISCOSITY_OK=FALSE per  | drop (PUB002)  |               |
|                    | becomes TRUE   | stays TRUE| PUB002                 |               |               |
+--------------------+----------------+----------+-------------------------+----------------+---------------+
*)

CASE BOOL_TO_INT(PASTE_E_STOP_NC) OF
    0: // Emergency stop active
        VFD_RUN := FALSE;
        ViscosityValid := FALSE;
        DebounceTimer(IN := FALSE, PT := DebounceTime);

    1: // Emergency stop cleared - normal operation
        IF NOT VISCOSITY_OK THEN
            ViscosityValid := FALSE;
            DebounceTimer(IN := FALSE, PT := DebounceTime);
        ELSE
            DebounceTimer(IN := TRUE, PT := DebounceTime);
            ViscosityValid := DebounceTimer.Q;
        END_IF;

        VFD_RUN := ViscosityValid;
END_CASE;

IF VFD_RUN THEN
    PUMP_RUNTIME_ACC := PUMP_RUNTIME_ACC + LTIME(CycleTime);
END_IF;

IF PUMP_RUNTIME_ACC >= tmp_MaintThreshold THEN
    PUMP_MAINT_DUE := TRUE;
END_IF;

END_FUNCTION_BLOCK

(* ---- public-easy-04.raw_candidate_02.st ---- *)
FUNCTION_BLOCK FB_JamPumpControl
VAR_INPUT
    VISCOSITY_OK    : BOOL;
    PASTE_E_STOP_NC : BOOL;
    DebounceTime    : TIME;
    CycleTime       : TIME;
END_VAR
VAR_OUTPUT
    VFD_RUN          : BOOL;
    PUMP_MAINT_DUE   : BOOL;
    PUMP_RUNTIME_ACC : LTIME;
END_VAR
VAR
    ViscosityValid : BOOL := FALSE;
    DebounceTimer  : TON;
    tmp_MaintThreshold : LTIME := LTIME#500h;
END_VAR

(* CONTRACT_RULES [] *)

(* ENGINEERING_CONTRACT
+====================+================+==========+=========================+================+===============+
| Output/State       | Activation     | Retention| Reset/Deactivation      | Same-Scan Prio | Boundaries    |
+====================+================+==========+=========================+================+===============+
| VFD_RUN            | ESTOP=TRUE     | Hold     | Immediately on ESTOP=FALSE per PUB003 | Immediate disable | Boolean       |
|                    | AND            |          | No delay on ESTOP loss   |               |               |
|                    | ViscosityValid |          |                          |               |               |
+--------------------+----------------+----------+-------------------------+----------------+---------------+
| ViscosityValid     | TON.Q=TRUE     | Hold TRUE| Invalidate on           | Immediate      | Internal state|
| (internal)         | after          | while    | VISCOSITY_OK=FALSE      | invalidation   |               |
|                    | DebounceTime   | VISCOSITY_OK=TRUE        | per PUB002     |               |               |
+--------------------+----------------+----------+-------------------------+----------------+---------------+
| PUMP_RUNTIME_ACC   | +CycleTime     | Preserve | Only via power-up init  | Increment per  | LTIME, max    |
|                    | per scan while | when     | (PUB006). No auto-reset | scan when      | 500h threshold|
|                    | VFD_RUN=TRUE   | stopped  | specified.              | VFD_RUN=TRUE   | for PUMP_MAINT|
+--------------------+----------------+----------+-------------------------+----------------+---------------+
| PUMP_MAINT_DUE     | Set when       | Hold TRUE| Not specified (informational per PUB005) | At threshold | Boolean       |
|                    | ACC >= 500h    |          | No reset required       |               |               |
+--------------------+----------------+----------+-------------------------+----------------+---------------+
| DebounceTimer      | Start when     | Running  | Reset (ET=TRUE) on      | Clear on input | TON; PT=DebounceTime |
|                    | VISCOSITY_OK   | if input | VISCOSITY_OK=FALSE per  | drop (PUB002)  |               |
|                    | becomes TRUE   | stays TRUE| PUB002                 |               |               |
+--------------------+----------------+----------+-------------------------+----------------+---------------+
*)

CASE BOOL_TO_INT(PASTE_E_STOP_NC) OF
    0: // Emergency stop active
        VFD_RUN := FALSE;
        ViscosityValid := FALSE;
        DebounceTimer(IN := FALSE, PT := DebounceTime);

    1: // Emergency stop cleared - normal operation
        IF NOT VISCOSITY_OK THEN
            ViscosityValid := FALSE;
            DebounceTimer(IN := FALSE, PT := DebounceTime);
        ELSE
            DebounceTimer(IN := TRUE, PT := DebounceTime);
            ViscosityValid := DebounceTimer.Q;
        END_IF;

        VFD_RUN := ViscosityValid;
END_CASE;

IF VFD_RUN THEN
    PUMP_RUNTIME_ACC := PUMP_RUNTIME_ACC + TIME_TO_LTIME(CycleTime);
END_IF;

IF PUMP_RUNTIME_ACC >= tmp_MaintThreshold THEN
    PUMP_MAINT_DUE := TRUE;
END_IF;

END_FUNCTION_BLOCK

(* ---- public-hard-03.candidate_01.st ---- *)
(* ENGINEERING_CONTRACT
| Output/State      | Activation          | Retention     | Reset               | Same-scan Priority | Units/Boundaries              |
|-------------------|---------------------|---------------|---------------------|--------------------|-------------------------------|
| recipeAdded       | addRecipe success   | Latched       | Implicit next call  | True               | status=16#0000 on success     |
| recipeDeleted     | deleteRecipe success| Latched       | Implicit next call  | True               | status=16#0000 on success     |
| recipeModified    | modifyRecipe success| Latched       | Implicit next call  | True               | status=16#0000 on success     |
| recipeQueryResult | queryRecipe found   | Held          | Implicit next call  | True               | Populated on match; preserved |
| error             | Any error condition | Latched       | Implicit next call  | True               | 16#8001-16#8005               |
| status            | Any operation       | Held          | Implicit next call  | True               | Error code or 0               |

Operation Order (same-scan priority): addRecipe > deleteRecipe > modifyRecipe > queryRecipe
Empty slot detection: recipeID = 0 in database slot
Duplicate detection: Any database slot with matching non-zero recipeID
Search scope: ARRAY[1..10] OF ST_Recipe, sequential scan
*)
(* CONTRACT_RULES [] *)

FUNCTION_BLOCK FB_RecipeManagement
VAR_INPUT
    addRecipe    : BOOL;
    deleteRecipe : BOOL;
    modifyRecipe : BOOL;
    queryRecipe  : BOOL;
    recipeIn     : ST_Recipe;
END_VAR
VAR_OUTPUT
    recipeAdded       : BOOL;
    recipeDeleted     : BOOL;
    recipeModified    : BOOL;
    recipeQueryResult : ST_Recipe;
    error             : BOOL;
    status            : WORD;
END_VAR
VAR_IN_OUT
    recipe : ARRAY[1..10] OF ST_Recipe;
END_VAR
VAR
    tmp_index     : INT;
    tmp_found     : BOOL;
    tmp_emptySlot : INT;
    tmp_emptyFound: BOOL;
END_VAR

    // Initialize outputs to safe state at start of scan
    recipeAdded  := FALSE;
    recipeDeleted  := FALSE;
    recipeModified := FALSE;
    error          := FALSE;
    status         := 16#0000;

    // Process operations in same-scan priority order: add > delete > modify > query
    // PUB010: Add Recipe
    IF addRecipe THEN
        tmp_found     := FALSE;
        tmp_emptySlot := 0;
        tmp_emptyFound := FALSE;
        tmp_index     := 1;

        // Search for duplicate and empty slot
        FOR tmp_index := 1 TO 10 DO
            IF recipe[tmp_index].recipeID = recipeIn.recipeID AND recipeIn.recipeID <> 0 THEN
                tmp_found := TRUE;
                EXIT;
            END_IF;
        END_FOR;

        IF NOT tmp_found THEN
            // No duplicate found, search for empty slot
            FOR tmp_index := 1 TO 10 DO
                IF recipe[tmp_index].recipeID = 0 THEN
                    tmp_emptySlot := tmp_index;
                    tmp_emptyFound := TRUE;
                    EXIT;
                END_IF;
            END_FOR;
        END_IF;

        IF tmp_found THEN
            // Duplicate recipe number exists
            // PUB010: error code 16#8002
            error  := TRUE;
            status := 16#8002;
        ELSIF NOT tmp_emptyFound THEN
            // No empty slot available
            // PUB010: error code 16#8003
            error  := TRUE;
            status := 16#8003;
        ELSE
            // Store in smallest index empty slot
            recipe[tmp_emptySlot] := recipeIn;
            recipeAdded := TRUE;
            error       := FALSE;
            status      := 16#0000;
        END_IF;
        RETURN;
    END_IF;

    // PUB011: Delete Recipe
    IF deleteRecipe THEN
        tmp_found := FALSE;
        tmp_index := 1;

        // Search for matching recipe number
        FOR tmp_index := 1 TO 10 DO
            IF recipe[tmp_index].recipeID = recipeIn.recipeID AND recipeIn.recipeID <> 0 THEN
                tmp_found := TRUE;
                EXIT;
            END_IF;
        END_FOR;

        IF NOT tmp_found THEN
            // Recipe number does not exist
            // PUB011: error code 16#8004
            error  := TRUE;
            status := 16#8004;
        ELSE
            // Delete recipe by setting recipeID to 0
            recipe[tmp_index].recipeID := 0;
            recipeDeleted := TRUE;
            error         := FALSE;
            status        := 16#0000;
        END_IF;
        RETURN;
    END_IF;

    // PUB012: Modify Recipe
    IF modifyRecipe THEN
        tmp_found := FALSE;
        tmp_index := 1;

        // Search for matching recipe number
        FOR tmp_index := 1 TO 10 DO
            IF recipe[tmp_index].recipeID = recipeIn.recipeID AND recipeIn.recipeID <> 0 THEN
                tmp_found := TRUE;
                EXIT;
            END_IF;
        END_FOR;

        IF NOT tmp_found THEN
            // Recipe number does not exist
            // PUB012: error code 16#8005
            error  := TRUE;
            status := 16#8005;
        ELSE
            // Replace recipe with input recipe
            recipe[tmp_index] := recipeIn;
            recipeModified := TRUE;
            error          := FALSE;
            status         := 16#0000;
        END_IF;
        RETURN;
    END_IF;

    // PUB009: Query Recipe
    IF queryRecipe THEN
        tmp_found := FALSE;
        tmp_index := 1;

        // Search for matching recipe number
        FOR tmp_index := 1 TO 10 DO
            IF recipe[tmp_index].recipeID = recipeIn.recipeID AND recipeIn.recipeID <> 0 THEN
                tmp_found := TRUE;
                recipeQueryResult := recipe[tmp_index];
                EXIT;
            END_IF;
        END_FOR;

        IF NOT tmp_found THEN
            // Recipe number does not exist
            // PUB009: error code 16#8001
            error  := TRUE;
            status := 16#8001;
        ELSE
            error  := FALSE;
            status := 16#0000;
        END_IF;
        RETURN;
    END_IF;

END_FUNCTION_BLOCK

(* ---- public-hard-03.candidate_02.st ---- *)
(* ENGINEERING_CONTRACT
| Output/State      | Activation          | Retention     | Reset               | Same-scan Priority | Units/Boundaries              |
|-------------------|---------------------|---------------|---------------------|--------------------|-------------------------------|
| recipeAdded       | addRecipe success   | Latched       | Implicit next call  | True               | status=16#0000 on success     |
| recipeDeleted     | deleteRecipe success| Latched       | Implicit next call  | True               | status=16#0000 on success     |
| recipeModified    | modifyRecipe success| Latched       | Implicit next call  | True               | status=16#0000 on success     |
| recipeQueryResult | queryRecipe found   | Held          | Implicit next call  | True               | Populated on match; preserved |
| error             | Any error condition | Latched       | Implicit next call  | True               | 16#8001-16#8005               |
| status            | Any operation       | Held          | Implicit next call  | True               | Error code or 0               |

Operation Order (same-scan priority): addRecipe > deleteRecipe > modifyRecipe > queryRecipe
Empty slot detection: recipeID = 0 in database slot
Duplicate detection: Any database slot with matching non-zero recipeID
Search scope: ARRAY[1..10] OF ST_Recipe, sequential scan
*)
(* CONTRACT_RULES [] *)

TYPE ST_Recipe :
STRUCT
    recipeID               : INT;
    ingredientType         : INT;
    ingredientRatio        : REAL;
    productionTemperature  : REAL;
END_STRUCT
END_TYPE;

FUNCTION_BLOCK FB_RecipeManagement
VAR_INPUT
    addRecipe    : BOOL;
    deleteRecipe : BOOL;
    modifyRecipe : BOOL;
    queryRecipe  : BOOL;
    recipeIn     : ST_Recipe;
END_VAR
VAR_OUTPUT
    recipeAdded       : BOOL;
    recipeDeleted     : BOOL;
    recipeModified    : BOOL;
    recipeQueryResult : ST_Recipe;
    error             : BOOL;
    status            : WORD;
END_VAR
VAR_IN_OUT
    recipe : ARRAY[1..10] OF ST_Recipe;
END_VAR
VAR
    tmp_index      : INT;
    tmp_found      : BOOL;
    tmp_emptySlot  : INT;
    tmp_emptyFound : BOOL;
END_VAR

    recipeAdded  := FALSE;
    recipeDeleted  := FALSE;
    recipeModified := FALSE;
    error          := FALSE;
    status         := 16#0000;

    IF addRecipe THEN
        tmp_found      := FALSE;
        tmp_emptySlot  := 0;
        tmp_emptyFound := FALSE;
        tmp_index      := 1;

        FOR tmp_index := 1 TO 10 DO
            IF recipe[tmp_index].recipeID = recipeIn.recipeID AND recipeIn.recipeID <> 0 THEN
                tmp_found := TRUE;
                EXIT;
            END_IF;
        END_FOR;

        IF NOT tmp_found THEN
            FOR tmp_index := 1 TO 10 DO
                IF recipe[tmp_index].recipeID = 0 THEN
                    tmp_emptySlot  := tmp_index;
                    tmp_emptyFound := TRUE;
                    EXIT;
                END_IF;
            END_FOR;
        END_IF;

        IF tmp_found THEN
            error  := TRUE;
            status := 16#8002;
        ELSIF NOT tmp_emptyFound THEN
            error  := TRUE;
            status := 16#8003;
        ELSE
            recipe[tmp_emptySlot] := recipeIn;
            recipeAdded := TRUE;
            error       := FALSE;
            status      := 16#0000;
        END_IF;
        RETURN;
    END_IF;

    IF deleteRecipe THEN
        tmp_found := FALSE;
        tmp_index := 1;

        FOR tmp_index := 1 TO 10 DO
            IF recipe[tmp_index].recipeID = recipeIn.recipeID AND recipeIn.recipeID <> 0 THEN
                tmp_found := TRUE;
                EXIT;
            END_IF;
        END_FOR;

        IF NOT tmp_found THEN
            error  := TRUE;
            status := 16#8004;
        ELSE
            recipe[tmp_index].recipeID := 0;
            recipeDeleted := TRUE;
            error         := FALSE;
            status        := 16#0000;
        END_IF;
        RETURN;
    END_IF;

    IF modifyRecipe THEN
        tmp_found := FALSE;
        tmp_index := 1;

        FOR tmp_index := 1 TO 10 DO
            IF recipe[tmp_index].recipeID = recipeIn.recipeID AND recipeIn.recipeID <> 0 THEN
                tmp_found := TRUE;
                EXIT;
            END_IF;
        END_FOR;

        IF NOT tmp_found THEN
            error  := TRUE;
            status := 16#8005;
        ELSE
            recipe[tmp_index] := recipeIn;
            recipeModified := TRUE;
            error          := FALSE;
            status         := 16#0000;
        END_IF;
        RETURN;
    END_IF;

    IF queryRecipe THEN
        tmp_found := FALSE;
        tmp_index := 1;

        FOR tmp_index := 1 TO 10 DO
            IF recipe[tmp_index].recipeID = recipeIn.recipeID AND recipeIn.recipeID <> 0 THEN
                tmp_found := TRUE;
                recipeQueryResult := recipe[tmp_index];
                EXIT;
            END_IF;
        END_FOR;

        IF NOT tmp_found THEN
            error  := TRUE;
            status := 16#8001;
        ELSE
            error  := FALSE;
            status := 16#0000;
        END_IF;
        RETURN;
    END_IF;

END_FUNCTION_BLOCK

(* ---- public-hard-03.candidate_03.st ---- *)
(* ENGINEERING_CONTRACT
| Output/State      | Activation          | Retention     | Reset               | Same-scan Priority | Units/Boundaries              |
|-------------------|---------------------|---------------|---------------------|--------------------|-------------------------------|
| recipeAdded       | addRecipe success   | Latched       | Implicit next call  | True               | status=16#0000 on success     |
| recipeDeleted     | deleteRecipe success| Latched       | Implicit next call  | True               | status=16#0000 on success     |
| recipeModified    | modifyRecipe success| Latched       | Implicit next call  | True               | status=16#0000 on success     |
| recipeQueryResult | queryRecipe found   | Held          | Implicit next call  | True               | Populated on match; preserved |
| error             | Any error condition | Latched       | Implicit next call  | True               | 16#8001-16#8005               |
| status            | Any operation       | Held          | Implicit next call  | True               | Error code or 0               |

Operation Order (same-scan priority): addRecipe > deleteRecipe > modifyRecipe > queryRecipe
Empty slot detection: recipeID = 0 in database slot
Duplicate detection: Any database slot with matching non-zero recipeID
Search scope: ARRAY[1..10] OF ST_Recipe, sequential scan
Bounded: status only changes when a command is processed; retained otherwise
*)
(* CONTRACT_RULES [] *)

TYPE ST_Recipe :
STRUCT
    recipeID               : INT;
    ingredientType         : INT;
    ingredientRatio        : REAL;
    productionTemperature  : REAL;
END_STRUCT
END_TYPE;

FUNCTION_BLOCK FB_RecipeManagement
VAR_INPUT
    addRecipe    : BOOL;
    deleteRecipe : BOOL;
    modifyRecipe : BOOL;
    queryRecipe  : BOOL;
    recipeIn     : ST_Recipe;
END_VAR
VAR_OUTPUT
    recipeAdded       : BOOL;
    recipeDeleted     : BOOL;
    recipeModified    : BOOL;
    recipeQueryResult : ST_Recipe;
    error             : BOOL;
    status            : WORD;
END_VAR
VAR_IN_OUT
    recipe : ARRAY[1..10] OF ST_Recipe;
END_VAR
VAR
    tmp_index      : INT;
    tmp_found      : BOOL;
    tmp_emptySlot  : INT;
    tmp_emptyFound : BOOL;
END_VAR

    recipeAdded  := FALSE;
    recipeDeleted  := FALSE;
    recipeModified := FALSE;

    IF addRecipe THEN
        tmp_found      := FALSE;
        tmp_emptySlot  := 0;
        tmp_emptyFound := FALSE;
        tmp_index      := 1;

        FOR tmp_index := 1 TO 10 DO
            IF recipe[tmp_index].recipeID = recipeIn.recipeID AND recipeIn.recipeID <> 0 THEN
                tmp_found := TRUE;
                EXIT;
            END_IF;
        END_FOR;

        IF tmp_found THEN
            error  := TRUE;
            status := 16#8002;
        ELSIF NOT tmp_emptyFound THEN
            error  := TRUE;
            status := 16#8003;
        ELSE
            recipe[tmp_emptySlot] := recipeIn;
            recipeAdded := TRUE;
            error       := FALSE;
            status      := 16#0000;
        END_IF;
        RETURN;
    END_IF;

    IF deleteRecipe THEN
        tmp_found := FALSE;
        tmp_index := 1;

        FOR tmp_index := 1 TO 10 DO
            IF recipe[tmp_index].recipeID = recipeIn.recipeID AND recipeIn.recipeID <> 0 THEN
                tmp_found := TRUE;
                EXIT;
            END_IF;
        END_FOR;

        IF NOT tmp_found THEN
            error  := TRUE;
            status := 16#8004;
        ELSE
            recipe[tmp_index].recipeID := 0;
            recipeDeleted := TRUE;
            error         := FALSE;
            status        := 16#0000;
        END_IF;
        RETURN;
    END_IF;

    IF modifyRecipe THEN
        tmp_found := FALSE;
        tmp_index := 1;

        FOR tmp_index := 1 TO 10 DO
            IF recipe[tmp_index].recipeID = recipeIn.recipeID AND recipeIn.recipeID <> 0 THEN
                tmp_found := TRUE;
                EXIT;
            END_IF;
        END_FOR;

        IF NOT tmp_found THEN
            error  := TRUE;
            status := 16#8005;
        ELSE
            recipe[tmp_index] := recipeIn;
            recipeModified := TRUE;
            error          := FALSE;
            status         := 16#0000;
        END_IF;
        RETURN;
    END_IF;

    IF queryRecipe THEN
        tmp_found := FALSE;
        tmp_index := 1;

        FOR tmp_index := 1 TO 10 DO
            IF recipe[tmp_index].recipeID = recipeIn.recipeID AND recipeIn.recipeID <> 0 THEN
                tmp_found := TRUE;
                recipeQueryResult := recipe[tmp_index];
                status := 16#0000;
                EXIT;
            END_IF;
        END_FOR;

        IF NOT tmp_found THEN
            error  := TRUE;
            status := 16#8001;
        END_IF;
        RETURN;
    END_IF;

END_FUNCTION_BLOCK

(* ---- public-hard-03.candidate_04.st ---- *)
Looking at the bounded status violations (S7, S9, S10 at position 2), the issue is that unconditional reset of `error` and `status` at the start of each call causes values to be cleared even when no operation is active. The bounded checker expects these values to persist between calls when no new operation is triggered, and to transition correctly through operation sequences.

The fix: Only reset `error` and `status` inside each active operation block, preserving state when no command input is asserted.

TYPE ST_Recipe :
STRUCT
    recipeID               : INT;
    ingredientType         : INT;
    ingredientRatio        : REAL;
    productionTemperature  : REAL;
END_STRUCT
END_TYPE

FUNCTION_BLOCK FB_RecipeManagement
VAR_INPUT
    addRecipe    : BOOL;
    deleteRecipe : BOOL;
    modifyRecipe : BOOL;
    queryRecipe  : BOOL;
    recipeIn     : ST_Recipe;
END_VAR
VAR_OUTPUT
    recipeAdded       : BOOL;
    recipeDeleted     : BOOL;
    recipeModified    : BOOL;
    recipeQueryResult : ST_Recipe;
    error             : BOOL;
    status            : WORD;
END_VAR
VAR_IN_OUT
    recipe : ARRAY[1..10] OF ST_Recipe;
END_VAR
VAR
    tmp_index      : INT;
    tmp_found      : BOOL;
    tmp_emptySlot  : INT;
    tmp_emptyFound : BOOL;
END_VAR

    recipeAdded  := FALSE;
    recipeDeleted  := FALSE;
    recipeModified := FALSE;

    IF addRecipe THEN
        error  := FALSE;
        status := 16#0000;

        tmp_found      := FALSE;
        tmp_emptySlot  := 0;
        tmp_emptyFound := FALSE;

        FOR tmp_index := 1 TO 10 DO
            IF recipe[tmp_index].recipeID = recipeIn.recipeID AND recipeIn.recipeID <> 0 THEN
                tmp_found := TRUE;
                EXIT;
            END_IF;
        END_FOR;

        IF NOT tmp_found THEN
            FOR tmp_index := 1 TO 10 DO
                IF recipe[tmp_index].recipeID = 0 THEN
                    tmp_emptySlot  := tmp_index;
                    tmp_emptyFound := TRUE;
                    EXIT;
                END_IF;
            END_FOR;
        END_IF;

        IF tmp_found THEN
            error  := TRUE;
            status := 16#8002;
        ELSIF NOT tmp_emptyFound THEN
            error  := TRUE;
            status := 16#8003;
        ELSE
            recipe[tmp_emptySlot] := recipeIn;
            recipeAdded := TRUE;
        END_IF;
        RETURN;
    END_IF;

    IF deleteRecipe THEN
        error  := FALSE;
        status := 16#0000;

        tmp_found := FALSE;

        FOR tmp_index := 1 TO 10 DO
            IF recipe[tmp_index].recipeID = recipeIn.recipeID AND recipeIn.recipeID <> 0 THEN
                tmp_found := TRUE;
                EXIT;
            END_IF;
        END_FOR;

        IF NOT tmp_found THEN
            error  := TRUE;
            status := 16#8004;
        ELSE
            recipe[tmp_index].recipeID := 0;
            recipeDeleted := TRUE;
        END_IF;
        RETURN;
    END_IF;

    IF modifyRecipe THEN
        error  := FALSE;
        status := 16#0000;

        tmp_found := FALSE;

        FOR tmp_index := 1 TO 10 DO
            IF recipe[tmp_index].recipeID = recipeIn.recipeID AND recipeIn.recipeID <> 0 THEN
                tmp_found := TRUE;
                EXIT;
            END_IF;
        END_FOR;

        IF NOT tmp_found THEN
            error  := TRUE;
            status := 16#8005;
        ELSE
            recipe[tmp_index] := recipeIn;
            recipeModified := TRUE;
        END_IF;
        RETURN;
    END_IF;

    IF queryRecipe THEN
        error  := FALSE;
        status := 16#0000;

        tmp_found := FALSE;

        FOR tmp_index := 1 TO 10 DO
            IF recipe[tmp_index].recipeID = recipeIn.recipeID AND recipeIn.recipeID <> 0 THEN
                tmp_found := TRUE;
                recipeQueryResult := recipe[tmp_index];
                EXIT;
            END_IF;
        END_FOR;

        IF NOT tmp_found THEN
            error  := TRUE;
            status := 16#8001;
        END_IF;
        RETURN;
    END_IF;

END_FUNCTION_BLOCK

(* ---- public-hard-03.raw_candidate_01.st ---- *)
(* ENGINEERING_CONTRACT
| Output/State      | Activation          | Retention     | Reset               | Same-scan Priority | Units/Boundaries              |
|-------------------|---------------------|---------------|---------------------|--------------------|-------------------------------|
| recipeAdded       | addRecipe success   | Latched       | Implicit next call  | True               | status=16#0000 on success     |
| recipeDeleted     | deleteRecipe success| Latched       | Implicit next call  | True               | status=16#0000 on success     |
| recipeModified    | modifyRecipe success| Latched       | Implicit next call  | True               | status=16#0000 on success     |
| recipeQueryResult | queryRecipe found   | Held          | Implicit next call  | True               | Populated on match; preserved |
| error             | Any error condition | Latched       | Implicit next call  | True               | 16#8001-16#8005               |
| status            | Any operation       | Held          | Implicit next call  | True               | Error code or 0               |

Operation Order (same-scan priority): addRecipe > deleteRecipe > modifyRecipe > queryRecipe
Empty slot detection: recipeID = 0 in database slot
Duplicate detection: Any database slot with matching non-zero recipeID
Search scope: ARRAY[1..10] OF ST_Recipe, sequential scan
*)
(* CONTRACT_RULES [] *)

FUNCTION_BLOCK FB_RecipeManagement
VAR_INPUT
    addRecipe    : BOOL;
    deleteRecipe : BOOL;
    modifyRecipe : BOOL;
    queryRecipe  : BOOL;
    recipeIn     : ST_Recipe;
END_VAR
VAR_OUTPUT
    recipeAdded       : BOOL;
    recipeDeleted     : BOOL;
    recipeModified    : BOOL;
    recipeQueryResult : ST_Recipe;
    error             : BOOL;
    status            : WORD;
END_VAR
VAR_IN_OUT
    recipe : ARRAY[1..10] OF ST_Recipe;
END_VAR
VAR
    tmp_index     : INT;
    tmp_found     : BOOL;
    tmp_emptySlot : INT;
    tmp_emptyFound: BOOL;
END_VAR

    // Initialize outputs to safe state at start of scan
    recipeAdded  := FALSE;
    recipeDeleted  := FALSE;
    recipeModified := FALSE;
    error          := FALSE;
    status         := 16#0000;

    // Process operations in same-scan priority order: add > delete > modify > query
    // PUB010: Add Recipe
    IF addRecipe THEN
        tmp_found     := FALSE;
        tmp_emptySlot := 0;
        tmp_emptyFound := FALSE;
        tmp_index     := 1;

        // Search for duplicate and empty slot
        FOR tmp_index := 1 TO 10 DO
            IF recipe[tmp_index].recipeID = recipeIn.recipeID AND recipeIn.recipeID <> 0 THEN
                tmp_found := TRUE;
                EXIT;
            END_IF
        END_FOR

        IF NOT tmp_found THEN
            // No duplicate found, search for empty slot
            FOR tmp_index := 1 TO 10 DO
                IF recipe[tmp_index].recipeID = 0 THEN
                    tmp_emptySlot := tmp_index;
                    tmp_emptyFound := TRUE;
                    EXIT;
                END_IF
            END_FOR
        END_IF

        IF tmp_found THEN
            // Duplicate recipe number exists
            // PUB010: error code 16#8002
            error  := TRUE;
            status := 16#8002;
        ELSIF NOT tmp_emptyFound THEN
            // No empty slot available
            // PUB010: error code 16#8003
            error  := TRUE;
            status := 16#8003;
        ELSE
            // Store in smallest index empty slot
            recipe[tmp_emptySlot] := recipeIn;
            recipeAdded := TRUE;
            error       := FALSE;
            status      := 16#0000;
        END_IF
        RETURN;
    END_IF

    // PUB011: Delete Recipe
    IF deleteRecipe THEN
        tmp_found := FALSE;
        tmp_index := 1;

        // Search for matching recipe number
        FOR tmp_index := 1 TO 10 DO
            IF recipe[tmp_index].recipeID = recipeIn.recipeID AND recipeIn.recipeID <> 0 THEN
                tmp_found := TRUE;
                EXIT;
            END_IF
        END_FOR

        IF NOT tmp_found THEN
            // Recipe number does not exist
            // PUB011: error code 16#8004
            error  := TRUE;
            status := 16#8004;
        ELSE
            // Delete recipe by setting recipeID to 0
            recipe[tmp_index].recipeID := 0;
            recipeDeleted := TRUE;
            error         := FALSE;
            status        := 16#0000;
        END_IF
        RETURN;
    END_IF

    // PUB012: Modify Recipe
    IF modifyRecipe THEN
        tmp_found := FALSE;
        tmp_index := 1;

        // Search for matching recipe number
        FOR tmp_index := 1 TO 10 DO
            IF recipe[tmp_index].recipeID = recipeIn.recipeID AND recipeIn.recipeID <> 0 THEN
                tmp_found := TRUE;
                EXIT;
            END_IF
        END_FOR

        IF NOT tmp_found THEN
            // Recipe number does not exist
            // PUB012: error code 16#8005
            error  := TRUE;
            status := 16#8005;
        ELSE
            // Replace recipe with input recipe
            recipe[tmp_index] := recipeIn;
            recipeModified := TRUE;
            error          := FALSE;
            status         := 16#0000;
        END_IF
        RETURN;
    END_IF

    // PUB009: Query Recipe
    IF queryRecipe THEN
        tmp_found := FALSE;
        tmp_index := 1;

        // Search for matching recipe number
        FOR tmp_index := 1 TO 10 DO
            IF recipe[tmp_index].recipeID = recipeIn.recipeID AND recipeIn.recipeID <> 0 THEN
                tmp_found := TRUE;
                recipeQueryResult := recipe[tmp_index];
                EXIT;
            END_IF
        END_FOR

        IF NOT tmp_found THEN
            // Recipe number does not exist
            // PUB009: error code 16#8001
            error  := TRUE;
            status := 16#8001;
        ELSE
            error  := FALSE;
            status := 16#0000;
        END_IF
        RETURN;
    END_IF

END_FUNCTION_BLOCK

(* ---- public-hard-03.raw_candidate_02.st ---- *)
(* ENGINEERING_CONTRACT
| Output/State      | Activation          | Retention     | Reset               | Same-scan Priority | Units/Boundaries              |
|-------------------|---------------------|---------------|---------------------|--------------------|-------------------------------|
| recipeAdded       | addRecipe success   | Latched       | Implicit next call  | True               | status=16#0000 on success     |
| recipeDeleted     | deleteRecipe success| Latched       | Implicit next call  | True               | status=16#0000 on success     |
| recipeModified    | modifyRecipe success| Latched       | Implicit next call  | True               | status=16#0000 on success     |
| recipeQueryResult | queryRecipe found   | Held          | Implicit next call  | True               | Populated on match; preserved |
| error             | Any error condition | Latched       | Implicit next call  | True               | 16#8001-16#8005               |
| status            | Any operation       | Held          | Implicit next call  | True               | Error code or 0               |

Operation Order (same-scan priority): addRecipe > deleteRecipe > modifyRecipe > queryRecipe
Empty slot detection: recipeID = 0 in database slot
Duplicate detection: Any database slot with matching non-zero recipeID
Search scope: ARRAY[1..10] OF ST_Recipe, sequential scan
*)
(* CONTRACT_RULES [] *)

TYPE ST_Recipe :
STRUCT
    recipeID               : INT;
    ingredientType         : INT;
    ingredientRatio        : REAL;
    productionTemperature  : REAL;
END_STRUCT
END_TYPE

FUNCTION_BLOCK FB_RecipeManagement
VAR_INPUT
    addRecipe    : BOOL;
    deleteRecipe : BOOL;
    modifyRecipe : BOOL;
    queryRecipe  : BOOL;
    recipeIn     : ST_Recipe;
END_VAR
VAR_OUTPUT
    recipeAdded       : BOOL;
    recipeDeleted     : BOOL;
    recipeModified    : BOOL;
    recipeQueryResult : ST_Recipe;
    error             : BOOL;
    status            : WORD;
END_VAR
VAR_IN_OUT
    recipe : ARRAY[1..10] OF ST_Recipe;
END_VAR
VAR
    tmp_index      : INT;
    tmp_found      : BOOL;
    tmp_emptySlot  : INT;
    tmp_emptyFound : BOOL;
END_VAR

    recipeAdded  := FALSE;
    recipeDeleted  := FALSE;
    recipeModified := FALSE;
    error          := FALSE;
    status         := 16#0000;

    IF addRecipe THEN
        tmp_found      := FALSE;
        tmp_emptySlot  := 0;
        tmp_emptyFound := FALSE;
        tmp_index      := 1;

        FOR tmp_index := 1 TO 10 DO
            IF recipe[tmp_index].recipeID = recipeIn.recipeID AND recipeIn.recipeID <> 0 THEN
                tmp_found := TRUE;
                EXIT;
            END_IF;
        END_FOR;

        IF NOT tmp_found THEN
            FOR tmp_index := 1 TO 10 DO
                IF recipe[tmp_index].recipeID = 0 THEN
                    tmp_emptySlot  := tmp_index;
                    tmp_emptyFound := TRUE;
                    EXIT;
                END_IF;
            END_FOR;
        END_IF;

        IF tmp_found THEN
            error  := TRUE;
            status := 16#8002;
        ELSIF NOT tmp_emptyFound THEN
            error  := TRUE;
            status := 16#8003;
        ELSE
            recipe[tmp_emptySlot] := recipeIn;
            recipeAdded := TRUE;
            error       := FALSE;
            status      := 16#0000;
        END_IF;
        RETURN;
    END_IF;

    IF deleteRecipe THEN
        tmp_found := FALSE;
        tmp_index := 1;

        FOR tmp_index := 1 TO 10 DO
            IF recipe[tmp_index].recipeID = recipeIn.recipeID AND recipeIn.recipeID <> 0 THEN
                tmp_found := TRUE;
                EXIT;
            END_IF;
        END_FOR;

        IF NOT tmp_found THEN
            error  := TRUE;
            status := 16#8004;
        ELSE
            recipe[tmp_index].recipeID := 0;
            recipeDeleted := TRUE;
            error         := FALSE;
            status        := 16#0000;
        END_IF;
        RETURN;
    END_IF;

    IF modifyRecipe THEN
        tmp_found := FALSE;
        tmp_index := 1;

        FOR tmp_index := 1 TO 10 DO
            IF recipe[tmp_index].recipeID = recipeIn.recipeID AND recipeIn.recipeID <> 0 THEN
                tmp_found := TRUE;
                EXIT;
            END_IF;
        END_FOR;

        IF NOT tmp_found THEN
            error  := TRUE;
            status := 16#8005;
        ELSE
            recipe[tmp_index] := recipeIn;
            recipeModified := TRUE;
            error          := FALSE;
            status         := 16#0000;
        END_IF;
        RETURN;
    END_IF;

    IF queryRecipe THEN
        tmp_found := FALSE;
        tmp_index := 1;

        FOR tmp_index := 1 TO 10 DO
            IF recipe[tmp_index].recipeID = recipeIn.recipeID AND recipeIn.recipeID <> 0 THEN
                tmp_found := TRUE;
                recipeQueryResult := recipe[tmp_index];
                EXIT;
            END_IF;
        END_FOR;

        IF NOT tmp_found THEN
            error  := TRUE;
            status := 16#8001;
        ELSE
            error  := FALSE;
            status := 16#0000;
        END_IF;
        RETURN;
    END_IF;

END_FUNCTION_BLOCK

(* ---- public-hard-03.raw_candidate_03.st ---- *)
(* ENGINEERING_CONTRACT
| Output/State      | Activation          | Retention     | Reset               | Same-scan Priority | Units/Boundaries              |
|-------------------|---------------------|---------------|---------------------|--------------------|-------------------------------|
| recipeAdded       | addRecipe success   | Latched       | Implicit next call  | True               | status=16#0000 on success     |
| recipeDeleted     | deleteRecipe success| Latched       | Implicit next call  | True               | status=16#0000 on success     |
| recipeModified    | modifyRecipe success| Latched       | Implicit next call  | True               | status=16#0000 on success     |
| recipeQueryResult | queryRecipe found   | Held          | Implicit next call  | True               | Populated on match; preserved |
| error             | Any error condition | Latched       | Implicit next call  | True               | 16#8001-16#8005               |
| status            | Any operation       | Held          | Implicit next call  | True               | Error code or 0               |

Operation Order (same-scan priority): addRecipe > deleteRecipe > modifyRecipe > queryRecipe
Empty slot detection: recipeID = 0 in database slot
Duplicate detection: Any database slot with matching non-zero recipeID
Search scope: ARRAY[1..10] OF ST_Recipe, sequential scan
Bounded: status only changes when a command is processed; retained otherwise
*)
(* CONTRACT_RULES [] *)

TYPE ST_Recipe :
STRUCT
    recipeID               : INT;
    ingredientType         : INT;
    ingredientRatio        : REAL;
    productionTemperature  : REAL;
END_STRUCT
END_TYPE;

FUNCTION_BLOCK FB_RecipeManagement
VAR_INPUT
    addRecipe    : BOOL;
    deleteRecipe : BOOL;
    modifyRecipe : BOOL;
    queryRecipe  : BOOL;
    recipeIn     : ST_Recipe;
END_VAR
VAR_OUTPUT
    recipeAdded       : BOOL;
    recipeDeleted     : BOOL;
    recipeModified    : BOOL;
    recipeQueryResult : ST_Recipe;
    error             : BOOL;
    status            : WORD;
END_VAR
VAR_IN_OUT
    recipe : ARRAY[1..10] OF ST_Recipe;
END_VAR
VAR
    tmp_index      : INT;
    tmp_found      : BOOL;
    tmp_emptySlot  : INT;
    tmp_emptyFound : BOOL;
END_VAR

    recipeAdded  := FALSE;
    recipeDeleted  := FALSE;
    recipeModified := FALSE;

    IF addRecipe THEN
        tmp_found      := FALSE;
        tmp_emptySlot  := 0;
        tmp_emptyFound := FALSE;
        tmp_index      := 1;

        FOR tmp_index := 1 TO 10 DO
            IF recipe[tmp_index].recipeID = recipeIn.recipeID AND recipeIn.recipeID <> 0 THEN
                tmp_found := TRUE;
                EXIT;
            END_IF;
        END_FOR;

        IF tmp_found THEN
            error  := TRUE;
            status := 16#8002;
        ELSIF NOT tmp_emptyFound THEN
            error  := TRUE;
            status := 16#8003;
        ELSE
            recipe[tmp_emptySlot] := recipeIn;
            recipeAdded := TRUE;
            error       := FALSE;
            status      := 16#0000;
        END_IF;
        RETURN;
    END_IF;

    IF deleteRecipe THEN
        tmp_found := FALSE;
        tmp_index := 1;

        FOR tmp_index := 1 TO 10 DO
            IF recipe[tmp_index].recipeID = recipeIn.recipeID AND recipeIn.recipeID <> 0 THEN
                tmp_found := TRUE;
                EXIT;
            END_IF;
        END_FOR;

        IF NOT tmp_found THEN
            error  := TRUE;
            status := 16#8004;
        ELSE
            recipe[tmp_index].recipeID := 0;
            recipeDeleted := TRUE;
            error         := FALSE;
            status        := 16#0000;
        END_IF;
        RETURN;
    END_IF;

    IF modifyRecipe THEN
        tmp_found := FALSE;
        tmp_index := 1;

        FOR tmp_index := 1 TO 10 DO
            IF recipe[tmp_index].recipeID = recipeIn.recipeID AND recipeIn.recipeID <> 0 THEN
                tmp_found := TRUE;
                EXIT;
            END_IF;
        END_FOR;

        IF NOT tmp_found THEN
            error  := TRUE;
            status := 16#8005;
        ELSE
            recipe[tmp_index] := recipeIn;
            recipeModified := TRUE;
            error          := FALSE;
            status         := 16#0000;
        END_IF;
        RETURN;
    END_IF;

    IF queryRecipe THEN
        tmp_found := FALSE;
        tmp_index := 1;

        FOR tmp_index := 1 TO 10 DO
            IF recipe[tmp_index].recipeID = recipeIn.recipeID AND recipeIn.recipeID <> 0 THEN
                tmp_found := TRUE;
                recipeQueryResult := recipe[tmp_index];
                status := 16#0000;
                EXIT;
            END_IF;
        END_FOR;

        IF NOT tmp_found THEN
            error  := TRUE;
            status := 16#8001;
        END_IF;
        RETURN;
    END_IF;

END_FUNCTION_BLOCK

(* ---- public-hard-03.raw_candidate_04.st ---- *)
Looking at the bounded status violations (S7, S9, S10 at position 2), the issue is that unconditional reset of `error` and `status` at the start of each call causes values to be cleared even when no operation is active. The bounded checker expects these values to persist between calls when no new operation is triggered, and to transition correctly through operation sequences.

The fix: Only reset `error` and `status` inside each active operation block, preserving state when no command input is asserted.

TYPE ST_Recipe :
STRUCT
    recipeID               : INT;
    ingredientType         : INT;
    ingredientRatio        : REAL;
    productionTemperature  : REAL;
END_STRUCT
END_TYPE

FUNCTION_BLOCK FB_RecipeManagement
VAR_INPUT
    addRecipe    : BOOL;
    deleteRecipe : BOOL;
    modifyRecipe : BOOL;
    queryRecipe  : BOOL;
    recipeIn     : ST_Recipe;
END_VAR
VAR_OUTPUT
    recipeAdded       : BOOL;
    recipeDeleted     : BOOL;
    recipeModified    : BOOL;
    recipeQueryResult : ST_Recipe;
    error             : BOOL;
    status            : WORD;
END_VAR
VAR_IN_OUT
    recipe : ARRAY[1..10] OF ST_Recipe;
END_VAR
VAR
    tmp_index      : INT;
    tmp_found      : BOOL;
    tmp_emptySlot  : INT;
    tmp_emptyFound : BOOL;
END_VAR

    recipeAdded  := FALSE;
    recipeDeleted  := FALSE;
    recipeModified := FALSE;

    IF addRecipe THEN
        error  := FALSE;
        status := 16#0000;

        tmp_found      := FALSE;
        tmp_emptySlot  := 0;
        tmp_emptyFound := FALSE;

        FOR tmp_index := 1 TO 10 DO
            IF recipe[tmp_index].recipeID = recipeIn.recipeID AND recipeIn.recipeID <> 0 THEN
                tmp_found := TRUE;
                EXIT;
            END_IF;
        END_FOR;

        IF NOT tmp_found THEN
            FOR tmp_index := 1 TO 10 DO
                IF recipe[tmp_index].recipeID = 0 THEN
                    tmp_emptySlot  := tmp_index;
                    tmp_emptyFound := TRUE;
                    EXIT;
                END_IF;
            END_FOR;
        END_IF;

        IF tmp_found THEN
            error  := TRUE;
            status := 16#8002;
        ELSIF NOT tmp_emptyFound THEN
            error  := TRUE;
            status := 16#8003;
        ELSE
            recipe[tmp_emptySlot] := recipeIn;
            recipeAdded := TRUE;
        END_IF;
        RETURN;
    END_IF;

    IF deleteRecipe THEN
        error  := FALSE;
        status := 16#0000;

        tmp_found := FALSE;

        FOR tmp_index := 1 TO 10 DO
            IF recipe[tmp_index].recipeID = recipeIn.recipeID AND recipeIn.recipeID <> 0 THEN
                tmp_found := TRUE;
                EXIT;
            END_IF;
        END_FOR;

        IF NOT tmp_found THEN
            error  := TRUE;
            status := 16#8004;
        ELSE
            recipe[tmp_index].recipeID := 0;
            recipeDeleted := TRUE;
        END_IF;
        RETURN;
    END_IF;

    IF modifyRecipe THEN
        error  := FALSE;
        status := 16#0000;

        tmp_found := FALSE;

        FOR tmp_index := 1 TO 10 DO
            IF recipe[tmp_index].recipeID = recipeIn.recipeID AND recipeIn.recipeID <> 0 THEN
                tmp_found := TRUE;
                EXIT;
            END_IF;
        END_FOR;

        IF NOT tmp_found THEN
            error  := TRUE;
            status := 16#8005;
        ELSE
            recipe[tmp_index] := recipeIn;
            recipeModified := TRUE;
        END_IF;
        RETURN;
    END_IF;

    IF queryRecipe THEN
        error  := FALSE;
        status := 16#0000;

        tmp_found := FALSE;

        FOR tmp_index := 1 TO 10 DO
            IF recipe[tmp_index].recipeID = recipeIn.recipeID AND recipeIn.recipeID <> 0 THEN
                tmp_found := TRUE;
                recipeQueryResult := recipe[tmp_index];
                EXIT;
            END_IF;
        END_FOR;

        IF NOT tmp_found THEN
            error  := TRUE;
            status := 16#8001;
        END_IF;
        RETURN;
    END_IF;

END_FUNCTION_BLOCK

(* ---- public-medium-03.candidate_01.st ---- *)
FUNCTION_BLOCK FB_MovingAverage
VAR_INPUT
    cyclicExecution : BOOL;
    trigger         : BOOL;
    value           : LREAL;
    windowSize      : INT;
    reset           : BOOL;
END_VAR

VAR_OUTPUT
    average           : LREAL;
    windowSizeReached : BOOL;
    error             : BOOL;
    status            : WORD;
END_VAR

VAR
    dataBuffer    : ARRAY[1..100] OF LREAL;
    currentIndex  : INT := 0;
    sampleCount   : INT := 0;
    sum           : LREAL := 0.0;
    tmp_lastTrigger : BOOL := FALSE;
END_VAR

(*
ENGINEERING_CONTRACT
===================
Operation Modes:
- cyclicExecution=TRUE: Update every scan cycle; trigger ignored (PUB002)
- cyclicExecution=FALSE: Rising edge on trigger updates average (PUB003)
- reset=TRUE: Clear all state, outputs to default, status=SUCCESS (PUB004)

Output Retention Policy:
| Output             | Activation         | Retention    | Reset by reset=TRUE |
|--------------------|--------------------|--------------|---------------------|
| average            | Each valid sample  | Hold last    | Yes (→0.0)          |
| windowSizeReached  | sampleCount>=winSz | Hold TRUE    | Yes (→FALSE)        |
| error              | windowSize<1 or >100| Hold TRUE   | Yes (→FALSE)        |
| status             | Per validation     | Hold code    | Yes (→SUCCESS)      |

Boundary Conditions:
- windowSize<1 OR >100 → error=TRUE, status=16#8200, skip processing (PUB004, PUB007)
- reset asserted → immediate clear, no processing (PUB004)
- Empty window (sampleCount=0) → average=0.0 (division-safe)
- Circular buffer wraps at windowSize, never exceeds 100 elements

Same-Scan Priority:
1. reset check (highest)
2. windowSize validation
3. trigger rising-edge detection
4. cyclicExecution evaluation
5. sample insertion / buffer rotation
6. average recalculation

Units: LREAL for all arithmetic (PUB001). windowSize in slots [1..100].
*)

(* CONTRACT_RULES
[
  {"kind": "hold_until_reset", "output": "windowSizeReached", "set_input": null, "reset_input": "reset"},
  {"kind": "hold_until_reset", "output": "error", "set_input": null, "reset_input": "reset"},
  {"kind": "hold_until_reset", "output": "status", "set_input": null, "reset_input": "reset"}
]
*)

    // Reset: clear all state and outputs
    IF reset THEN
        currentIndex     := 0;
        sampleCount      := 0;
        sum              := 0.0;
        average          := 0.0;
        windowSizeReached := FALSE;
        error            := FALSE;
        status           := 16#0000;
        tmp_lastTrigger  := FALSE;
        RETURN;
    END_IF;

    // Validate window size (PUB007)
    IF windowSize < 1 OR windowSize > 100 THEN
        error  := TRUE;
        status := 16#8200;
        RETURN;
    END_IF;

    // No validation error; set success status (PUB006)
    error  := FALSE;
    status := 16#0000;

    // Determine if a new sample should be processed (PUB002, PUB003)
    tmp_newSample := FALSE;
    IF cyclicExecution THEN
        tmp_newSample := TRUE;
    ELSIF trigger AND NOT tmp_lastTrigger THEN
        tmp_newSample := TRUE;
    END_IF;
    tmp_lastTrigger := trigger;

    // Process new data point if triggered (PUB001)
    IF tmp_newSample THEN
        // Clamp effective window to array upper bound (100)
        tmp_effectiveWindow := windowSize;
        IF tmp_effectiveWindow > 100 THEN
            tmp_effectiveWindow := 100;
        END_IF;

        IF sampleCount < tmp_effectiveWindow THEN
            // Window not yet full: append new value
            sampleCount := sampleCount + 1;
            dataBuffer[sampleCount] := value;
            sum := sum + value;
        ELSE
            // Window full: rotate out oldest value using circular buffer
            currentIndex := (currentIndex MOD tmp_effectiveWindow) + 1;
            sum := sum - dataBuffer[currentIndex] + value;
            dataBuffer[currentIndex] := value;
        END_IF;
    END_IF;

    // Calculate moving arithmetic mean (PUB001)
    IF sampleCount > 0 THEN
        average := sum / TO_LREAL(sampleCount);
    ELSE
        average := 0.0;
    END_IF;

    // Indicate whether maximum window width has been reached (PUB001)
    tmp_effectiveWindow := windowSize;
    IF tmp_effectiveWindow > 100 THEN
        tmp_effectiveWindow := 100;
    END_IF;
    windowSizeReached := (sampleCount >= tmp_effectiveWindow);

END_FUNCTION_BLOCK
